// TIA Portal V20 export
// export: Created 2026-10-20T12:52:55.7604709Z, ExportSetting WithDefaults, DisplayName Totally Integrated Automation Portal, DisplayVersion V20 Update 6, DisplayName TIA Portal Openness, DisplayVersion V20 Update 6, DisplayName TIA Portal Version Control Interface, DisplayVersion V20 Update 6, DisplayName SINAMICS Startdrive Advanced, DisplayVersion V20 SP1, DisplayName SINAMICS Startdrive G130, G150, S120, S150, SINAMICS MV, G220, S200, S210, DisplayVersion V20 SP1, DisplayName SINAMICS Startdrive G110M, G120, G120C, G120D, G120P, G115D, DisplayVersion V20 SP1, DisplayName STEP 7 Professional, DisplayVersion V20 Update 6, DisplayName STEP 7 Safety, DisplayVersion V20 Update 2, DisplayName WinCC Basic/Comfort/Advanced, DisplayVersion V20 Update 6, DisplayName WinCC Unified, DisplayVersion V20 Update 6
DATA_BLOCK "DB_Receive_Data_From_Logistex"   // DB900
{ S7_Optimized_Access := 'TRUE' }
VERSION : 0.1
// stored: AutoNumber false, DBAccessibleFromOPCUA true, IsOnlyStoredInLoadMemory false, IsRetainMemResEnabled false, IsWriteProtectedInAS false, MemoryReserve 100
   VAR
      J1310_Conv_Infeed : "Conv_Infeed";
      J1320_Conv_Infeed { S7_SetPoint := 'True'} : "Conv_Infeed";
      J1330_Conv_Infeed { S7_SetPoint := 'True'} : "Conv_Infeed";
      J1310_Conv_Oufeed { S7_SetPoint := 'True'} : "Conv_Outfeed";
      J1320_Conv_Oufeed { S7_SetPoint := 'True'} : "Conv_Outfeed";
      J1330_Conv_Oufeed { S7_SetPoint := 'True'} : "Conv_Outfeed";
      CNV_STATUS : Array[1..10] of Byte;
      PLC_STATUS : Struct
         Hardbit : Bool;
         "PLC_E-Stop" : Bool;
      END_STRUCT;
   END_VAR
BEGIN
END_DATA_BLOCK
